// TIA Portal V20 export
// export: Created 2026-10-19T18:35:58.3200796Z, ExportSetting WithDefaults, DisplayName Totally Integrated Automation Portal, DisplayVersion V20 Update 6, DisplayName TIA Portal Openness, DisplayVersion V20 Update 6, DisplayName TIA Portal Version Control Interface, DisplayVersion V20 Update 6, DisplayName SINAMICS Startdrive Advanced, DisplayVersion V20 SP1, DisplayName SINAMICS Startdrive G130, G150, S120, S150, SINAMICS MV, G220, S200, S210, DisplayVersion V20 SP1, DisplayName SINAMICS Startdrive G110M, G120, G120C, G120D, G120P, G115D, DisplayVersion V20 SP1, DisplayName STEP 7 Professional, DisplayVersion V20 Update 6, DisplayName STEP 7 Safety, DisplayVersion V20 Update 2, DisplayName WinCC Basic/Comfort/Advanced, DisplayVersion V20 Update 6, DisplayName WinCC Unified, DisplayVersion V20 Update 6
DATA_BLOCK "Force"   // DB12
{ S7_Optimized_Access := 'TRUE' }
VERSION : 0.1
// stored: AutoNumber true, DBAccessibleFromOPCUA true, IsOnlyStoredInLoadMemory false, IsRetainMemResEnabled false, IsWriteProtectedInAS false, MemoryReserve 100
   VAR
      Remote_Panel : Array[1..2] of Struct
         "CX101_SFTY STOPPER ROTATE" : Bool;
         "CX102_SFTY STOPPER ROTATE" : Bool;
         "CX103_SFTY STOPPER ROTATE" : Bool;
         "CX104_SFTY STOPPER ROTATE" : Bool;
         "CX105_SFTY STOPPER ROTATE" : Bool;
         "CX106_SFTY STOPPER ROTATE" : Bool;
         "CX107_SFTY STOPPER ROTATE" : Bool;
         "CX108_SFTY STOPPER ROTATE" : Bool;
         "VTDx DOCKING PINS 1 RETRACT" : Bool;
         "VTDx DOCKING PINS 1 EXTEND" : Bool;
         "VTDx DOCKING PINS 2 EXTEND" : Bool;
         "VTDx DOCKING PINS 2 RETRACT" : Bool;
         "SCA X00Y STACK LIGHTS ORANGE" : Bool;
         "SCA X00Y STACK LIGHTS GREEN" : Bool;
         "SCA X00Y STACK LIGHTS RED" : Bool;
         "EMERGENCY STOP RESET STATUS - ON(X)" : Bool;
      END_STRUCT;
   END_VAR
BEGIN
END_DATA_BLOCK
